// TIA Portal V20 export
// export: Created 2026-10-12T05:42:35.9235091Z, ExportSetting WithDefaults, DisplayName Totally Integrated Automation Portal, DisplayVersion V20, DisplayName TIA Portal Openness, DisplayVersion V20, DisplayName TIA Portal Teamcenter Gateway, DisplayVersion V20, DisplayName TIA Portal Version Control Interface, DisplayVersion V20, DisplayName SINAMICS Startdrive Advanced, DisplayVersion V20 SP1 Update 2, DisplayName SINAMICS Startdrive G110M, G120, G120C, G120D, G120P, G115D, DisplayVersion V20 SP1 Update 2, DisplayName SINAMICS Startdrive G130, G150, S120, S150, SINAMICS MV, G220, S200, S210, DisplayVersion V20 SP1 Update 2, DisplayName STEP 7 Professional, DisplayVersion V20, DisplayName STEP 7 Safety, DisplayVersion V20, DisplayName WinCC Basic/Comfort/Advanced, DisplayVersion V20, DisplayName WinCC Professional, DisplayVersion V20, DisplayName WinCC Unified, DisplayVersion V20
FUNCTION_BLOCK "FB_PressDemoHardwareDriver"   // FB14, SCL
{ S7_Optimized_Access := 'TRUE' }
VERSION : 0.1
// stored: AutoNumber true, IsIECCheckEnabled false, IsRetainMemResEnabled false, MemoryReserve 100, SetENOAutomatically false, UDAEnableTagReadback false
   VAR_INPUT
      ReadInputs { ExternalAccessible := 'False'; ExternalVisible := 'False'; ExternalWritable := 'False'} : Bool;
   END_VAR
BEGIN

   IF #ReadInputs THEN
       "GDB_FraktalHal".Data.PressDemo.Process.PartPresent := "GDB_PressDemoIO".PartPresent;
       "GDB_FraktalHal".Data.PressDemo.Process.PartQuality := "GDB_PressDemoIO".PartQuality;
       "GDB_FraktalHal".Data.PressDemo.Process.AirPressureOk := "GDB_PressDemoIO".AirPressureOk;
       "GDB_FraktalHal".Data.PressDemo.Process.TwoHandHeld := "GDB_PressDemoIO".TwoHandHeld;
       "GDB_FraktalHal".Data.PressDemo.Process.StartPulse := "GDB_PressDemoIO".StartPulse;
       "GDB_FraktalHal".Data.PressDemo.PressRam.FeedbackExtended := "GDB_PressDemoIO".RamExtended;
       "GDB_FraktalHal".Data.PressDemo.PressRam.FeedbackRetracted := "GDB_PressDemoIO".RamRetracted;
       "GDB_FraktalHal".Data.PressDemo.Door.FeedbackExtended := "GDB_PressDemoIO".DoorClosed;
       "GDB_FraktalHal".Data.PressDemo.Door.FeedbackRetracted := "GDB_PressDemoIO".DoorOpen;
       "GDB_FraktalHal".Data.PressDemo.PartSlide.FeedbackExtended := "GDB_PressDemoIO".SlideInside;
       "GDB_FraktalHal".Data.PressDemo.PartSlide.FeedbackRetracted := "GDB_PressDemoIO".SlideOutside;
   ELSE
       "GDB_PressDemoIO".RamExtend := "GDB_FraktalHal".Data.PressDemo.PressRam.CoilExtend;
       "GDB_PressDemoIO".RamRetract := "GDB_FraktalHal".Data.PressDemo.PressRam.CoilRetract;
       "GDB_PressDemoIO".DoorClose := "GDB_FraktalHal".Data.PressDemo.Door.CoilExtend;
       "GDB_PressDemoIO".DoorRelease := "GDB_FraktalHal".Data.PressDemo.Door.CoilRetract;
       "GDB_PressDemoIO".SlideExtend := "GDB_FraktalHal".Data.PressDemo.PartSlide.CoilExtend;
       "GDB_PressDemoIO".SlideRetract := "GDB_FraktalHal".Data.PressDemo.PartSlide.CoilRetract;
   END_IF;
END_FUNCTION_BLOCK
